(* IEC 61131-3 sources: volt/packages/volt-lsp-iec/test-corpus/twincat-project14/TwinCAT Project14/PLC/Untitled2/Untitled2 Project/References/Tc2_Standard, 32 files *)

(* ---- Global_Version.gvl ---- *)
VAR_GLOBAL
	stLibVersion_Tc2_Standard : ST_LibVersion;
END_VAR

(* ---- CONCAT.pou ---- *)
FUNCTION CONCAT : STRING(255)
VAR_INPUT
	STR1 : STRING(255);
	STR2 : STRING(255);
END_VAR
END_FUNCTION

(* ---- DELETE.pou ---- *)
FUNCTION DELETE : STRING(255)
VAR_INPUT
	STR : STRING(255);
	LEN : INT;
	POS : INT;
END_VAR
END_FUNCTION

(* ---- FIND.pou ---- *)
FUNCTION FIND : INT
VAR_INPUT
	STR1 : STRING(255);
	STR2 : STRING(255);
END_VAR
END_FUNCTION

(* ---- INSERT.pou ---- *)
FUNCTION INSERT : STRING(255)
VAR_INPUT
	STR1 : STRING(255);
	STR2 : STRING(255);
	POS : INT;
END_VAR
END_FUNCTION

(* ---- LEFT.pou ---- *)
FUNCTION LEFT : STRING(255)
VAR_INPUT
	STR : STRING(255);
	SIZE : INT;
END_VAR
END_FUNCTION

(* ---- LEN.pou ---- *)
FUNCTION LEN : INT
VAR_INPUT
	STR : STRING(255);
END_VAR
END_FUNCTION

(* ---- MID.pou ---- *)
FUNCTION MID : STRING(255)
VAR_INPUT
	STR : STRING(255);
	LEN : INT;
	POS : INT;
END_VAR
END_FUNCTION

(* ---- REPLACE.pou ---- *)
FUNCTION REPLACE : STRING(255)
VAR_INPUT
	STR1 : STRING(255);
	STR2 : STRING(255);
	L : INT;
	P : INT;
END_VAR
END_FUNCTION

(* ---- RIGHT.pou ---- *)
FUNCTION RIGHT : STRING(255)
VAR_INPUT
	STR : STRING(255);
	SIZE : INT;
END_VAR
END_FUNCTION

(* ---- WCONCAT.pou ---- *)
FUNCTION WCONCAT : WSTRING(255)
VAR_INPUT
	STR1 : WSTRING(255);
	STR2 : WSTRING(255);
END_VAR
END_FUNCTION

(* ---- WDELETE.pou ---- *)
FUNCTION WDELETE : WSTRING(255)
VAR_INPUT
	STR : WSTRING(255);
	LEN : INT;
	POS : INT;
END_VAR
END_FUNCTION

(* ---- WFIND.pou ---- *)
FUNCTION WFIND : INT
VAR_INPUT
	STR1 : WSTRING(255);
	STR2 : WSTRING(255);
END_VAR
END_FUNCTION

(* ---- WINSERT.pou ---- *)
FUNCTION WINSERT : WSTRING(255)
VAR_INPUT
	STR1 : WSTRING(255);
	STR2 : WSTRING(255);
	POS : INT;
END_VAR
END_FUNCTION

(* ---- WLEFT.pou ---- *)
FUNCTION WLEFT : WSTRING(255)
VAR_INPUT
	STR : WSTRING(255);
	SIZE : INT;
END_VAR
END_FUNCTION

(* ---- WLEN.pou ---- *)
FUNCTION WLEN : INT
VAR_INPUT
	STR : WSTRING(255);
END_VAR
END_FUNCTION

(* ---- WMID.pou ---- *)
FUNCTION WMID : WSTRING(255)
VAR_INPUT
	STR : WSTRING(255);
	LEN : INT;
	POS : INT;
END_VAR
END_FUNCTION

(* ---- WREPLACE.pou ---- *)
FUNCTION WREPLACE : WSTRING(255)
VAR_INPUT
	STR1 : WSTRING(255);
	STR2 : WSTRING(255);
	L : INT;
	P : INT;
END_VAR
END_FUNCTION

(* ---- WRIGHT.pou ---- *)
FUNCTION WRIGHT : WSTRING(255)
VAR_INPUT
	STR : WSTRING(255);
	SIZE : INT;
END_VAR
END_FUNCTION

(* ---- CTD.pou ---- *)
FUNCTION_BLOCK CTD
VAR_INPUT
	CD : BOOL;
	LOAD : BOOL;
	PV : WORD;
END_VAR
VAR_OUTPUT
	Q : BOOL;
	CV : WORD;
END_VAR
END_FUNCTION_BLOCK

(* ---- CTU.pou ---- *)
FUNCTION_BLOCK CTU
VAR_INPUT
	CU : BOOL;
	RESET : BOOL;
	PV : WORD;
END_VAR
VAR_OUTPUT
	Q : BOOL;
	CV : WORD;
END_VAR
END_FUNCTION_BLOCK

(* ---- CTUD.pou ---- *)
FUNCTION_BLOCK CTUD
VAR_INPUT
	CU : BOOL;
	CD : BOOL;
	RESET : BOOL;
	LOAD : BOOL;
	PV : WORD;
END_VAR
VAR_OUTPUT
	QU : BOOL;
	QD : BOOL;
	CV : WORD;
END_VAR
END_FUNCTION_BLOCK

(* ---- F_TRIG.pou ---- *)
FUNCTION_BLOCK F_TRIG
VAR_INPUT
	CLK : BOOL;
END_VAR
VAR_OUTPUT
	Q : BOOL;
END_VAR
END_FUNCTION_BLOCK

(* ---- LTOF.pou ---- *)
FUNCTION_BLOCK LTOF
VAR_INPUT
	IN : BOOL;
	PT : LTIME;
END_VAR
VAR_OUTPUT
	Q : BOOL;
	ET : LTIME;
END_VAR
END_FUNCTION_BLOCK

(* ---- LTON.pou ---- *)
FUNCTION_BLOCK LTON
VAR_INPUT
	IN : BOOL;
	PT : LTIME;
END_VAR
VAR_OUTPUT
	Q : BOOL;
	ET : LTIME;
END_VAR
END_FUNCTION_BLOCK

(* ---- LTP.pou ---- *)
FUNCTION_BLOCK LTP
VAR_INPUT
	IN : BOOL;
	PT : LTIME;
END_VAR
VAR_OUTPUT
	Q : BOOL;
	ET : LTIME;
END_VAR
END_FUNCTION_BLOCK

(* ---- R_TRIG.pou ---- *)
FUNCTION_BLOCK R_TRIG
VAR_INPUT
	CLK : BOOL;
END_VAR
VAR_OUTPUT
	Q : BOOL;
END_VAR
END_FUNCTION_BLOCK

(* ---- RS.pou ---- *)
FUNCTION_BLOCK RS
VAR_INPUT
	SET : BOOL;
	RESET1 : BOOL;
END_VAR
VAR_OUTPUT
	Q1 : BOOL;
END_VAR
END_FUNCTION_BLOCK

(* ---- SR.pou ---- *)
FUNCTION_BLOCK SR
VAR_INPUT
	SET1 : BOOL;
	RESET : BOOL;
END_VAR
VAR_OUTPUT
	Q1 : BOOL;
END_VAR
END_FUNCTION_BLOCK

(* ---- TOF.pou ---- *)
FUNCTION_BLOCK TOF
VAR_INPUT
	IN : BOOL;
	PT : TIME;
END_VAR
VAR_OUTPUT
	Q : BOOL;
	ET : TIME;
END_VAR
END_FUNCTION_BLOCK

(* ---- TON.pou ---- *)
FUNCTION_BLOCK TON
VAR_INPUT
	IN : BOOL;
	PT : TIME;
END_VAR
VAR_OUTPUT
	Q : BOOL;
	ET : TIME;
END_VAR
END_FUNCTION_BLOCK

(* ---- TP.pou ---- *)
FUNCTION_BLOCK TP
VAR_INPUT
	IN : BOOL;
	PT : TIME;
END_VAR
VAR_OUTPUT
	Q : BOOL;
	ET : TIME;
END_VAR
END_FUNCTION_BLOCK
